SUBAPPLICATION Dauerfunktion (* Subapplication Type *)
  (* Standard: 61499-2 *)
  (* Version 1.0, 2023-01-29, Franz *)
  IMPORT DefaultPool::SoftKey_Licht;
  IMPORT isobus::UT::io::Softkey::SoftKeyActivationCode::SK_RELEASED;
  IMPORT DefaultPool::AuxInput_Licht;
  IMPORT isobus::UT::io::Auxiliary::IN::AuxiliaryState::AuxDisabled;
  IMPORT DataPanel::io::MI::DQ::DataPanel_MI_DO::DigitalOutput_8A;
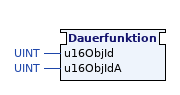
  VAR_INPUT
    u16ObjId : UINT;
    u16ObjIdA : UINT;
  END_VAR
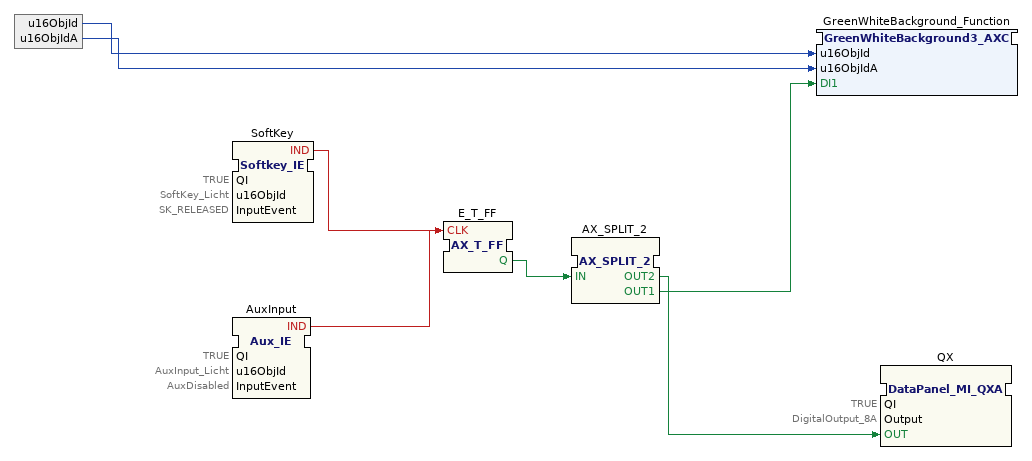
  FBS
    E_T_FF : adapter::events::unidirectional::AX_T_FF;
    QX : DataPanel::io::MI::DQ::DataPanel_MI_QXA(QI := TRUE, Output := DigitalOutput_8A);
    SoftKey : isobus::UT::io::Softkey::Softkey_IE(QI := TRUE, u16ObjId := SoftKey_Licht, InputEvent := SK_RELEASED);
    AuxInput : isobus::UT::io::Auxiliary::IN::Aux_IE(QI := TRUE, u16ObjId := AuxInput_Licht, InputEvent := AuxDisabled);
    AX_SPLIT_2 : adapter::events::unidirectional::AX_SPLIT_2;
  END_FBS
  SUBAPPS
    GreenWhiteBackground_Function : MyLib::sys::GreenWhiteBackground3_AXC;
  END_SUBAPPS
  EVENT_CONNECTIONS
    SoftKey.IND TO E_T_FF.CLK;
    AuxInput.IND TO E_T_FF.CLK;
  END_CONNECTIONS
  DATA_CONNECTIONS
    u16ObjId TO GreenWhiteBackground_Function.u16ObjId;
    u16ObjIdA TO GreenWhiteBackground_Function.u16ObjIdA;
  END_CONNECTIONS
  ADAPTER_CONNECTIONS
    AX_SPLIT_2.OUT2 TO QX.OUT;
    E_T_FF.Q TO AX_SPLIT_2.IN;
    AX_SPLIT_2.OUT1 TO GreenWhiteBackground_Function.DI1;
  END_CONNECTIONS
END_SUBAPPLICATION
